SUBAPPLICATION NumericValue_TO_AUI2_AND_STORE_PUBLISH (* Kopie von NumericValue_TO_AUI2_AND_STORE, zusaetzlich mit M2M-Publish des bestaetigten Werts (AUI_SPLIT_2 -> AUI_SPLIT_3: 3. Zweig fuer AUI_PUBLISH_1). Der M2M-Publish haengt damit am selben, bereits bewaehrten internen Confirm-Rueckpfad wie VT-Anzeige (AUI_TO_AUDI) und INI-Persistenz (INI_AUI) - kein fragiler externer Selfloop auf einem zusaetzlichen AUI2_TO_AUI-Bruecken- Baustein mehr noetig, der bei einem externen Umbau vergessen werden kann (Franz, nach Live-Debug einer genau solchen Regression: 'eine Kopie machen, und der PUBLISH kommt da innen rein'). *)
  (* Standard: 61499-2; Description: Copyright (c) 2026 Büngener Schuder GmbH This program and the accompanying materials are made available under the terms of the Eclipse Public License 2.0 which is available at https://www.eclipse.org/legal/epl-2.0/ SPDX-License-Identifier: EPL-2.0 *)
  (* Version 1.1, 2026-11-13, Franz Höpfinger, Meisterschulen am Ostbahnhof, Neuer Eingang DEFAULT_VALUE (bisher fest 0) an INI_AUI.DEFAULT_VALUE - je Instanz einstellbar, Default unveraendert 0. *)
  (* Version 1.0, 2026-10-14, Franz Höpfinger, Büngener Schuder GmbH, initial implementation - Kopie von NumericValue_TO_AUI2_AND_STORE v3.0, AUI_SPLIT_2 zu AUI_SPLIT_3 erweitert, neuer InputVar ID_WRITE + AUI_PUBLISH_1 (M2M) am 3. Split-Ausgang. Erster Aufrufer: BunkerKlappen_Fanghaken_Option.SUB (ersetzt den externen AUI2_TO_AUI+Selfloop+AUI_SPLIT_2 fuer den M2M-Pfad, der heute per Regression gebrochen war - der verbleibende externe AUI2_TO_AUI dort wird nur noch fuer den rein lokalen DEMUX-Tap gebraucht). *)
  PACKAGE MyLib::sys;
  IMPORT isobus::UT::Q::const::IDs::ID_NULL;
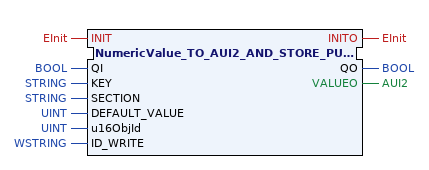
  EVENT_INPUT
    INIT : EInit; (* Initialization Request *)
  END_EVENT
  EVENT_OUTPUT
    INITO : EInit; (* Initialization Confirm *)
  END_EVENT
  VAR_INPUT
    QI : BOOL := TRUE; (* Quality Input - TRUE to enable service *)
    KEY : STRING; (* Key name. *)
    SECTION : STRING; (* Section name. *)
    DEFAULT_VALUE : UINT := UINT#0; (* Wert, wenn der KEY noch nicht in der INI steht *)
    u16ObjId : UINT := ID_NULL; (* Object ID *)
    ID_WRITE : WSTRING; (* Lokale Publish-Adresse (ACTION=WRITE) fuer den bestaetigten Wert - M2M, wird remote abonniert *)
  END_VAR
  VAR_OUTPUT
    QO : BOOL; (* Quality Output - TRUE if service executed successfully *)
  END_VAR
  PLUGS
    VALUEO : adapter::types::bidirectional::AUI2;
  END_PLUGS
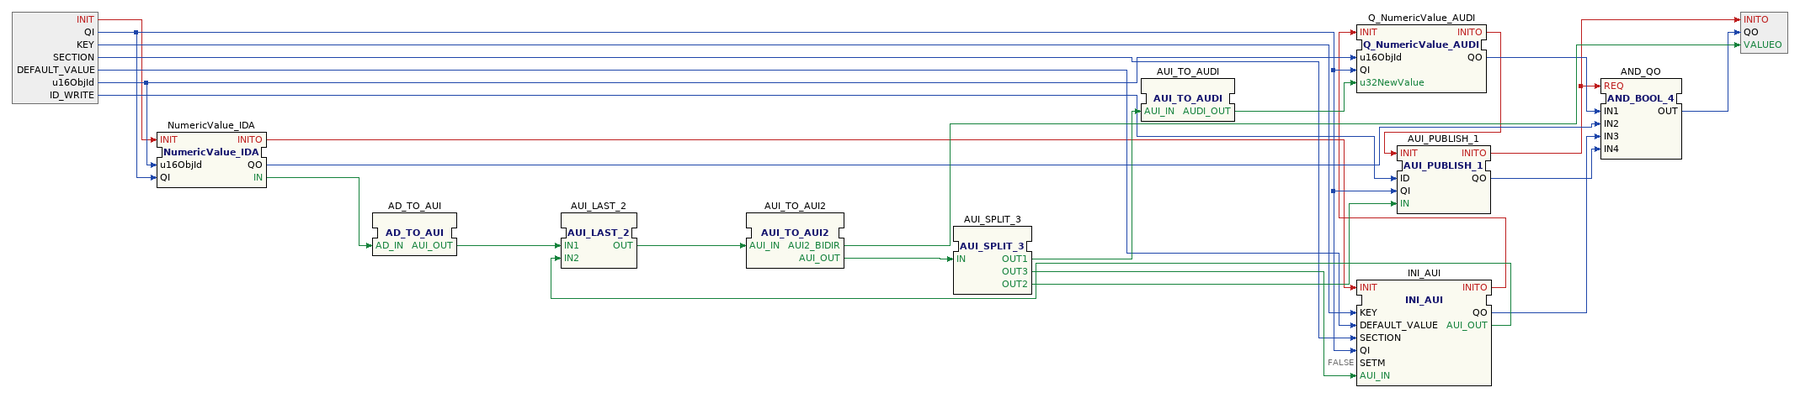
  (* SETM=FALSE: INI_AUI2 quittiert nur beim Boot (INIT->INITO->GET->GETO) automatisch, NICHT bei jedem spaeteren Schreibvorgang ueber VAL (Vorwaertsrichtung). Der Boot-Wert laeuft ueber AUI_TO_AUI2_1.AUI_OUT zu AUI_LAST_2 (siehe oben) und gewinnt dort einmalig gegen die Live-VT-Lesung. Waere SETM=TRUE, wuerde jeder spaetere Schreibvorgang sofort ein neues Echo auf AUI_OUT ausloesen, das wieder bei AUI_LAST_2 ankaeme und erneut Richtung VALUEO geschickt wuerde - ein Dauerkreislauf. *)
  FBS
    NumericValue_IDA : isobus::UT::io::NumericValue::NumericValue_IDA;
    AD_TO_AUI : adapter::conversion::unidirectional::AD_TO_AUI;
    AUI_TO_AUI2 : adapter::conversion::bidirectional::AUI_TO_AUI2; (* Bruecke zum externen Consumer (z.B. AOption_AUI_DEMUX_N.K) *)
    AUI_TO_AUDI : adapter::conversion::unidirectional::AUI_TO_AUDI;
    Q_NumericValue_AUDI : isobus::UT::Q::Q_NumericValue_AUDI;
    AUI_LAST_2 : adapter::events::unidirectional::AUI_LAST_2; (* Last-Writer-Wins: beim Boot gewinnt der INI_AUI2-Wert (IN2), danach jede Live-VT-Aenderung (IN1) *)
    AUI_SPLIT_3 : adapter::events::unidirectional::AUI_SPLIT_3; (* 3. Zweig (OUT3) fuer AUI_PUBLISH_1 - der bestaetigte Wert (aus AUI_TO_AUI2.AUI_OUT) wird jetzt auch direkt M2M published, am selben Confirm-Rueckpfad wie VT-Anzeige/INI-Persistenz *)
    INI_AUI : eclipse4diac::storage::INI_AUI(SETM := FALSE);
    AUI_PUBLISH_1 : adapter::net::AUI_PUBLISH_1;
    AND_QO : iec61131::booleanOperators::AND_BOOL_4;
  END_FBS
  EVENT_CONNECTIONS
    INIT TO NumericValue_IDA.INIT;
    NumericValue_IDA.INITO TO INI_AUI.INIT;
    INI_AUI.INITO TO Q_NumericValue_AUDI.INIT;
    Q_NumericValue_AUDI.INITO TO AUI_PUBLISH_1.INIT;
    AUI_PUBLISH_1.INITO TO INITO;
    AUI_PUBLISH_1.INITO TO AND_QO.REQ;
  END_CONNECTIONS
  DATA_CONNECTIONS
    KEY TO INI_AUI.KEY;
    DEFAULT_VALUE TO INI_AUI.DEFAULT_VALUE;
    SECTION TO INI_AUI.SECTION;
    u16ObjId TO NumericValue_IDA.u16ObjId;
    u16ObjId TO Q_NumericValue_AUDI.u16ObjId;
    ID_WRITE TO AUI_PUBLISH_1.ID;
    QI TO Q_NumericValue_AUDI.QI;
    QI TO NumericValue_IDA.QI;
    QI TO INI_AUI.QI;
    QI TO AUI_PUBLISH_1.QI;
    Q_NumericValue_AUDI.QO TO AND_QO.IN1;
    NumericValue_IDA.QO TO AND_QO.IN2;
    INI_AUI.QO TO AND_QO.IN3;
    AUI_PUBLISH_1.QO TO AND_QO.IN4;
    AND_QO.OUT TO QO;
  END_CONNECTIONS
  ADAPTER_CONNECTIONS
    NumericValue_IDA.IN TO AD_TO_AUI.AD_IN;
    AD_TO_AUI.AUI_OUT TO AUI_LAST_2.IN1;
    AUI_LAST_2.OUT TO AUI_TO_AUI2.AUI_IN;
    AUI_TO_AUI2.AUI2_BIDIR TO VALUEO;
    AUI_TO_AUDI.AUDI_OUT TO Q_NumericValue_AUDI.u32NewValue;
    AUI_SPLIT_3.OUT1 TO AUI_TO_AUDI.AUI_IN;
    AUI_SPLIT_3.OUT3 TO INI_AUI.AUI_IN;
    INI_AUI.AUI_OUT TO AUI_LAST_2.IN2;
    AUI_TO_AUI2.AUI_OUT TO AUI_SPLIT_3.IN;
    AUI_SPLIT_3.OUT2 TO AUI_PUBLISH_1.IN;
  END_CONNECTIONS
END_SUBAPPLICATION
